(* IEC 61131-3 sources: trust-platform/crates/trust-runtime/tests/fixtures/plcopen_motion/homing_negative_deferred_public_surface/src, 2 files *)

(* ---- main.st ---- *)
VAR_GLOBAL
    g_trust_motion_axis_initialized : ARRAY[0..31] OF BOOL;
    g_trust_motion_state : ARRAY[0..31] OF MC_AXIS_STATUS;
    g_trust_motion_grouped : ARRAY[0..31] OF BOOL;
    g_trust_motion_power_command : ARRAY[0..31] OF BOOL;
    g_trust_motion_power_stage : ARRAY[0..31] OF BOOL;
    g_trust_motion_axis_error : ARRAY[0..31] OF WORD;
    g_trust_motion_actual_position : ARRAY[0..31] OF REAL;
    g_trust_motion_set_position : ARRAY[0..31] OF REAL;
    g_trust_motion_commanded_position : ARRAY[0..31] OF REAL;
    g_trust_motion_actual_velocity : ARRAY[0..31] OF REAL;
    g_trust_motion_set_velocity : ARRAY[0..31] OF REAL;
    g_trust_motion_commanded_velocity : ARRAY[0..31] OF REAL;
    g_trust_motion_actual_torque : ARRAY[0..31] OF REAL;
    g_trust_motion_home_abs_switch : ARRAY[0..31] OF BOOL;
    g_trust_motion_limit_switch_pos : ARRAY[0..31] OF BOOL;
    g_trust_motion_limit_switch_neg : ARRAY[0..31] OF BOOL;
    g_trust_motion_simulation : ARRAY[0..31] OF BOOL;
    g_trust_motion_communication_ready : ARRAY[0..31] OF BOOL;
    g_trust_motion_ready_for_power_on : ARRAY[0..31] OF BOOL;
    g_trust_motion_is_homed : ARRAY[0..31] OF BOOL;
    g_trust_motion_axis_warning : ARRAY[0..31] OF BOOL;
    g_trust_motion_constant_velocity : ARRAY[0..31] OF BOOL;
    g_trust_motion_accelerating : ARRAY[0..31] OF BOOL;
    g_trust_motion_decelerating : ARRAY[0..31] OF BOOL;
    g_trust_motion_vel_factor : ARRAY[0..31] OF REAL;
    g_trust_motion_acc_factor : ARRAY[0..31] OF REAL;
    g_trust_motion_jerk_factor : ARRAY[0..31] OF REAL;
    g_trust_motion_sw_limit_pos : ARRAY[0..31] OF REAL;
    g_trust_motion_sw_limit_neg : ARRAY[0..31] OF REAL;
    g_trust_motion_enable_limit_pos : ARRAY[0..31] OF BOOL;
    g_trust_motion_enable_limit_neg : ARRAY[0..31] OF BOOL;
    g_trust_motion_enable_pos_lag_monitoring : ARRAY[0..31] OF BOOL;
    g_trust_motion_max_position_lag : ARRAY[0..31] OF REAL;
    g_trust_motion_max_velocity_system : ARRAY[0..31] OF REAL;
    g_trust_motion_max_velocity_appl : ARRAY[0..31] OF REAL;
    g_trust_motion_max_acceleration_system : ARRAY[0..31] OF REAL;
    g_trust_motion_max_acceleration_appl : ARRAY[0..31] OF REAL;
    g_trust_motion_max_deceleration_system : ARRAY[0..31] OF REAL;
    g_trust_motion_max_deceleration_appl : ARRAY[0..31] OF REAL;
    g_trust_motion_max_jerk_system : ARRAY[0..31] OF REAL;
    g_trust_motion_max_jerk_appl : ARRAY[0..31] OF REAL;
    g_trust_motion_resolved_acceleration : ARRAY[0..31] OF REAL;
    g_trust_motion_resolved_deceleration : ARRAY[0..31] OF REAL;
    g_trust_motion_resolved_jerk : ARRAY[0..31] OF REAL;
    g_trust_motion_next_command_id : ARRAY[0..31] OF UINT;
    g_trust_motion_active_command_id : ARRAY[0..31] OF UINT;
    g_trust_motion_active_command_kind : ARRAY[0..31] OF TRUST_MOTION_COMMAND_KIND;
    g_trust_motion_active_buffer_mode : ARRAY[0..31] OF MC_BUFFER_MODE;
    g_trust_motion_queue_depth : ARRAY[0..31] OF UINT;
    g_trust_motion_queue0_command_id : ARRAY[0..31] OF UINT;
    g_trust_motion_queue0_command_kind : ARRAY[0..31] OF TRUST_MOTION_COMMAND_KIND;
    g_trust_motion_queue0_buffer_mode : ARRAY[0..31] OF MC_BUFFER_MODE;
    g_trust_motion_queue1_command_id : ARRAY[0..31] OF UINT;
    g_trust_motion_queue1_command_kind : ARRAY[0..31] OF TRUST_MOTION_COMMAND_KIND;
    g_trust_motion_queue1_buffer_mode : ARRAY[0..31] OF MC_BUFFER_MODE;
    g_trust_motion_aborted0_command_id : ARRAY[0..31] OF UINT;
    g_trust_motion_aborted1_command_id : ARRAY[0..31] OF UINT;
    g_trust_motion_aborted2_command_id : ARRAY[0..31] OF UINT;
    g_trust_motion_vendor_bool_1000 : ARRAY[0..31] OF BOOL;
    g_trust_motion_ref_signal_active : ARRAY[0..31] OF BOOL;
    g_trust_motion_ref_signal_position : ARRAY[0..31] OF REAL;
    g_trust_motion_ref_signal_code : ARRAY[0..31] OF UINT;
    g_trust_motion_abs_encoder_position : ARRAY[0..31] OF REAL;
    g_trust_motion_distance_coded_ready : ARRAY[0..31] OF BOOL;
    g_trust_motion_distance_coded_position : ARRAY[0..31] OF REAL;
END_VAR

PROGRAM Main
END_PROGRAM

(* ---- tests.st ---- *)
PROGRAM plcopen_motion_homing_deferred_public_surface_is_absent
VAR
    StepReferenceFlyingSwitch : MC_StepReferenceFlyingSwitch;
    StepReferenceFlyingRefPulse : MC_StepReferenceFlyingRefPulse;
    AbortPassiveHoming : MC_AbortPassiveHoming;
END_VAR
END_PROGRAM
